RoboDK station: Doosan_M0609_SSM3_Experiment.rdk

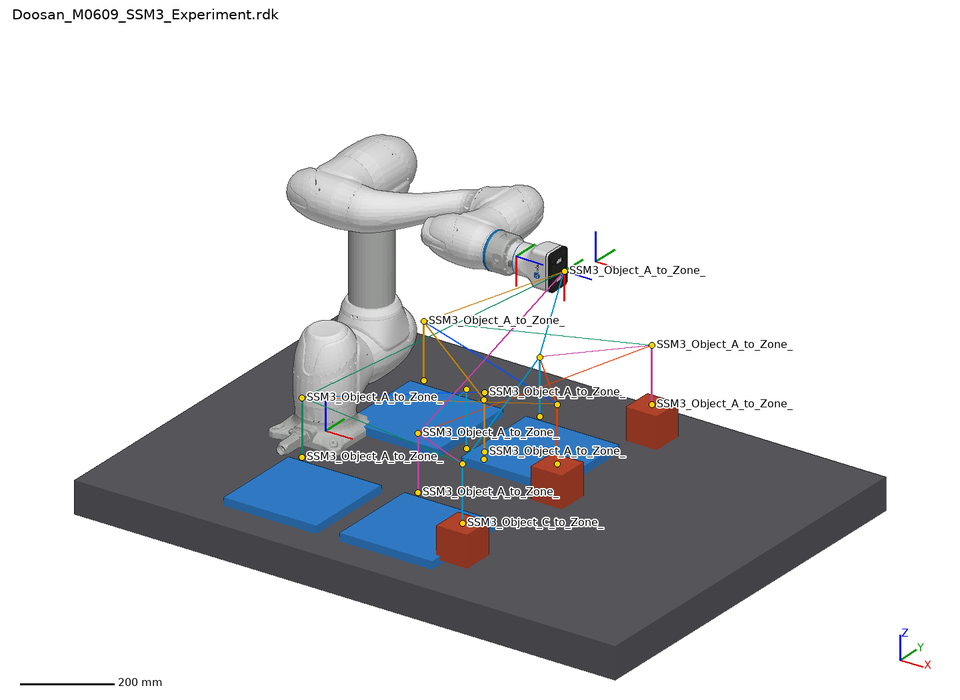
[picture v0: the station drawn from its stored meshes, robots at their saved joint values, targets as dots, program paths as lines]
Station Doosan_M0609_Pick_and_Place (saved by RoboDK 6.1.1). Poses are relative to the parent item; angles as X-Y-Z fixed-axis rotations.
  - frame Robot_Base at (0, 0, 0) mm
    - robot Doosan Robotics M0609 White: 6 axes, payload 6 kg, reach 900 mm, repeatability 0.03 mm, weight 27 kg
        modified DH rows (alpha deg, a mm, theta deg, d mm): 0, 0, 0, 135; -90, 0, -90, -6.207; 0, 411, -90, 0; -90, 0, 0, 368; 90, 0, 0, 0; -90, 0, 180, 121
        base shift (0, 0, 0) mm, rotated rx 0 ry 0 rz 180 deg
        joint limits [-360, -360, -150, -360, -360, -360] to [360, 360, 150, 360, 360, 360]; home [0, 0, 90, 0, 0, 0]; saved at [0, 0, 90, 0, 0, 0]
      - tool SSM3_Motion_TCP, TCP at (0, 0, 125) mm
      - frame OnRobot-2FG7-Gripper at (0, 0, 0) mm
        - robot OnRobot-2FG7-Gripper-Mechanism: 1 axes
            joint limits [0] to [55]; home [0]; saved at [49.5]
      - frame AUTO_Attach_TCP at (0, 0, 125) mm
  - frame TEST3 at (0, 1000, 0) mm
  - frame SSM3_Workcell at (0, 0, 0) mm
    - object SSM3_Table at (400, 0, -40) mm, size 1400 x 1000 x 80 mm, geometry from SSM3_Table.stl
    - object SSM3_Zone_A at (150, -300, 10) mm, size 240 x 240 x 20 mm, geometry from SSM3_Zone_A.stl
    - object SSM3_Zone_B at (450, -300, 10) mm, size 240 x 240 x 20 mm, geometry from SSM3_Zone_B.stl
    - object SSM3_Zone_C at (150, 150, 10) mm, size 240 x 240 x 20 mm, geometry from SSM3_Zone_C.stl
    - object SSM3_Zone_D at (450, 150, 10) mm, size 240 x 240 x 20 mm, geometry from SSM3_Zone_D.stl
    - target SSM3_Object_A_to_Zone_A_Home (Cartesian target) at (614, 6.21, 546) mm, rotated rx 0 ry 90 rz 0 deg; joints [0, 0, 90, 0, 0, 0] of Doosan Robotics M0609 White
    - target SSM3_Object_A_to_Zone_A_PickApproach (Cartesian target) at (440, -40, 230) mm, rotated rx 180 ry 0 rz 0 deg; joints [0, 0, 90, 0, 0, 0] of Doosan Robotics M0609 White
    - target SSM3_Object_A_to_Zone_A_Pick (Cartesian target) at (440, -40, 90) mm, rotated rx 180 ry 0 rz 0 deg; joints [0, 0, 90, 0, 0, 0] of Doosan Robotics M0609 White
    - target SSM3_Object_A_to_Zone_A_PlaceApproach (Cartesian target) at (150, -300, 240) mm, rotated rx 180 ry 0 rz 0 deg; joints [0, 0, 90, 0, 0, 0] of Doosan Robotics M0609 White
    - target SSM3_Object_A_to_Zone_A_Place (Cartesian target) at (150, -300, 100) mm, rotated rx 180 ry 0 rz 0 deg; joints [0, 0, 90, 0, 0, 0] of Doosan Robotics M0609 White
    - target SSM3_Object_A_to_Zone_B_Home (Cartesian target) at (614, 6.21, 546) mm, rotated rx 0 ry 90 rz 0 deg; joints [0, 0, 90, 0, 0, 0] of Doosan Robotics M0609 White
    - target SSM3_Object_A_to_Zone_B_PickApproach (Cartesian target) at (600, 350, 230) mm, rotated rx 180 ry 0 rz 0 deg; joints [0, 0, 90, 0, 0, 0] of Doosan Robotics M0609 White
    - target SSM3_Object_A_to_Zone_B_Pick (Cartesian target) at (600, 350, 90) mm, rotated rx 180 ry 0 rz 0 deg; joints [0, 0, 90, 0, 0, 0] of Doosan Robotics M0609 White
    - target SSM3_Object_A_to_Zone_B_PlaceApproach (Cartesian target) at (450, -300, 240) mm, rotated rx 180 ry 0 rz 0 deg; joints [0, 0, 90, 0, 0, 0] of Doosan Robotics M0609 White
    - target SSM3_Object_A_to_Zone_B_Place (Cartesian target) at (450, -300, 100) mm, rotated rx 180 ry 0 rz 0 deg; joints [0, 0, 90, 0, 0, 0] of Doosan Robotics M0609 White
    - target SSM3_Object_A_to_Zone_C_Home (Cartesian target) at (614, 6.21, 546) mm, rotated rx 0 ry 90 rz 0 deg; joints [0, 0, 90, 0, 0, 0] of Doosan Robotics M0609 White
    - target SSM3_Object_A_to_Zone_C_PickApproach (Cartesian target) at (600, 350, 230) mm, rotated rx 180 ry 0 rz 0 deg; joints [0, 0, 90, 0, 0, 0] of Doosan Robotics M0609 White
    - target SSM3_Object_A_to_Zone_C_Pick (Cartesian target) at (600, 350, 90) mm, rotated rx 180 ry 0 rz 0 deg; joints [0, 0, 90, 0, 0, 0] of Doosan Robotics M0609 White
    - target SSM3_Object_A_to_Zone_C_PlaceApproach (Cartesian target) at (150, 150, 240) mm, rotated rx 180 ry 0 rz 0 deg; joints [0, 0, 90, 0, 0, 0] of Doosan Robotics M0609 White
    - target SSM3_Object_A_to_Zone_C_Place (Cartesian target) at (150, 150, 100) mm, rotated rx 180 ry 0 rz 0 deg; joints [0, 0, 90, 0, 0, 0] of Doosan Robotics M0609 White
    - target SSM3_Object_A_to_Zone_D_Home (Cartesian target) at (614, 6.21, 546) mm, rotated rx 0 ry 90 rz 0 deg; joints [0, 0, 90, 0, 0, 0] of Doosan Robotics M0609 White
    - target SSM3_Object_A_to_Zone_D_PickApproach (Cartesian target) at (600, 350, 230) mm, rotated rx 180 ry 0 rz 0 deg; joints [0, 0, 90, 0, 0, 0] of Doosan Robotics M0609 White
    - target SSM3_Object_A_to_Zone_D_Pick (Cartesian target) at (600, 350, 90) mm, rotated rx 180 ry 0 rz 0 deg; joints [0, 0, 90, 0, 0, 0] of Doosan Robotics M0609 White
    - target SSM3_Object_A_to_Zone_D_PlaceApproach (Cartesian target) at (450, 150, 240) mm, rotated rx 180 ry 0 rz 0 deg; joints [0, 0, 90, 0, 0, 0] of Doosan Robotics M0609 White
    - target SSM3_Object_A_to_Zone_D_Place (Cartesian target) at (450, 150, 100) mm, rotated rx 180 ry 0 rz 0 deg; joints [0, 0, 90, 0, 0, 0] of Doosan Robotics M0609 White
    - target SSM3_Object_B_to_Zone_A_Home (Cartesian target) at (614, 6.21, 546) mm, rotated rx 0 ry 90 rz 0 deg; joints [0, 0, 90, 0, 0, 0] of Doosan Robotics M0609 White
    - target SSM3_Object_B_to_Zone_A_PickApproach (Cartesian target) at (600, 0, 230) mm, rotated rx 180 ry 0 rz 0 deg; joints [0, 0, 90, 0, 0, 0] of Doosan Robotics M0609 White
    - target SSM3_Object_B_to_Zone_A_Pick (Cartesian target) at (600, 0, 90) mm, rotated rx 180 ry 0 rz 0 deg; joints [0, 0, 90, 0, 0, 0] of Doosan Robotics M0609 White
    - target SSM3_Object_B_to_Zone_A_PlaceApproach (Cartesian target) at (150, -300, 240) mm, rotated rx 180 ry 0 rz 0 deg; joints [0, 0, 90, 0, 0, 0] of Doosan Robotics M0609 White
    - target SSM3_Object_B_to_Zone_A_Place (Cartesian target) at (150, -300, 100) mm, rotated rx 180 ry 0 rz 0 deg; joints [0, 0, 90, 0, 0, 0] of Doosan Robotics M0609 White
    - target SSM3_Object_B_to_Zone_B_Home (Cartesian target) at (614, 6.21, 546) mm, rotated rx 0 ry 90 rz 0 deg; joints [0, 0, 90, 0, 0, 0] of Doosan Robotics M0609 White
    - target SSM3_Object_B_to_Zone_B_PickApproach (Cartesian target) at (400, -50, 230) mm, rotated rx 180 ry 0 rz 0 deg; joints [0, 0, 90, 0, 0, 0] of Doosan Robotics M0609 White
    - target SSM3_Object_B_to_Zone_B_Pick (Cartesian target) at (400, -50, 90) mm, rotated rx 180 ry 0 rz 0 deg; joints [0, 0, 90, 0, 0, 0] of Doosan Robotics M0609 White
    - target SSM3_Object_B_to_Zone_B_PlaceApproach (Cartesian target) at (450, -300, 240) mm, rotated rx 180 ry 0 rz 0 deg; joints [0, 0, 90, 0, 0, 0] of Doosan Robotics M0609 White
    - target SSM3_Object_B_to_Zone_B_Place (Cartesian target) at (450, -300, 100) mm, rotated rx 180 ry 0 rz 0 deg; joints [0, 0, 90, 0, 0, 0] of Doosan Robotics M0609 White
    - target SSM3_Object_B_to_Zone_C_Home (Cartesian target) at (614, 6.21, 546) mm, rotated rx 0 ry 90 rz 0 deg; joints [0, 0, 90, 0, 0, 0] of Doosan Robotics M0609 White
    - target SSM3_Object_B_to_Zone_C_PickApproach (Cartesian target) at (600, 0, 230) mm, rotated rx 180 ry 0 rz 0 deg; joints [0, 0, 90, 0, 0, 0] of Doosan Robotics M0609 White
    - target SSM3_Object_B_to_Zone_C_Pick (Cartesian target) at (600, 0, 90) mm, rotated rx 180 ry 0 rz 0 deg; joints [0, 0, 90, 0, 0, 0] of Doosan Robotics M0609 White
    - target SSM3_Object_B_to_Zone_C_PlaceApproach (Cartesian target) at (150, 150, 240) mm, rotated rx 180 ry 0 rz 0 deg; joints [0, 0, 90, 0, 0, 0] of Doosan Robotics M0609 White
    - target SSM3_Object_B_to_Zone_C_Place (Cartesian target) at (150, 150, 100) mm, rotated rx 180 ry 0 rz 0 deg; joints [0, 0, 90, 0, 0, 0] of Doosan Robotics M0609 White
    - target SSM3_Object_B_to_Zone_D_Home (Cartesian target) at (614, 6.21, 546) mm, rotated rx 0 ry 90 rz 0 deg; joints [0, 0, 90, 0, 0, 0] of Doosan Robotics M0609 White
    - target SSM3_Object_B_to_Zone_D_PickApproach (Cartesian target) at (600, 0, 230) mm, rotated rx 180 ry 0 rz 0 deg; joints [0, 0, 90, 0, 0, 0] of Doosan Robotics M0609 White
    - target SSM3_Object_B_to_Zone_D_Pick (Cartesian target) at (600, 0, 90) mm, rotated rx 180 ry 0 rz 0 deg; joints [0, 0, 90, 0, 0, 0] of Doosan Robotics M0609 White
    - target SSM3_Object_B_to_Zone_D_PlaceApproach (Cartesian target) at (450, 150, 240) mm, rotated rx 180 ry 0 rz 0 deg; joints [0, 0, 90, 0, 0, 0] of Doosan Robotics M0609 White
    - target SSM3_Object_B_to_Zone_D_Place (Cartesian target) at (450, 150, 100) mm, rotated rx 180 ry 0 rz 0 deg; joints [0, 0, 90, 0, 0, 0] of Doosan Robotics M0609 White
    - target SSM3_Object_C_to_Zone_A_Home (Cartesian target) at (614, 6.21, 546) mm, rotated rx 0 ry 90 rz 0 deg; joints [0, 0, 90, 0, 0, 0] of Doosan Robotics M0609 White
    - target SSM3_Object_C_to_Zone_A_PickApproach (Cartesian target) at (600, -350, 230) mm, rotated rx 180 ry 0 rz 0 deg; joints [0, 0, 90, 0, 0, 0] of Doosan Robotics M0609 White
    - target SSM3_Object_C_to_Zone_A_Pick (Cartesian target) at (600, -350, 90) mm, rotated rx 180 ry 0 rz 0 deg; joints [0, 0, 90, 0, 0, 0] of Doosan Robotics M0609 White
    - target SSM3_Object_C_to_Zone_A_PlaceApproach (Cartesian target) at (150, -300, 240) mm, rotated rx 180 ry 0 rz 0 deg; joints [0, 0, 90, 0, 0, 0] of Doosan Robotics M0609 White
    - target SSM3_Object_C_to_Zone_A_Place (Cartesian target) at (150, -300, 100) mm, rotated rx 180 ry 0 rz 0 deg; joints [0, 0, 90, 0, 0, 0] of Doosan Robotics M0609 White
    - target SSM3_Object_C_to_Zone_B_Home (Cartesian target) at (614, 6.21, 546) mm, rotated rx 0 ry 90 rz 0 deg; joints [0, 0, 90, 0, 0, 0] of Doosan Robotics M0609 White
    - target SSM3_Object_C_to_Zone_B_PickApproach (Cartesian target) at (600, -350, 230) mm, rotated rx 180 ry 0 rz 0 deg; joints [0, 0, 90, 0, 0, 0] of Doosan Robotics M0609 White
    - target SSM3_Object_C_to_Zone_B_Pick (Cartesian target) at (600, -350, 90) mm, rotated rx 180 ry 0 rz 0 deg; joints [0, 0, 90, 0, 0, 0] of Doosan Robotics M0609 White
    - target SSM3_Object_C_to_Zone_B_PlaceApproach (Cartesian target) at (450, -300, 240) mm, rotated rx 180 ry 0 rz 0 deg; joints [0, 0, 90, 0, 0, 0] of Doosan Robotics M0609 White
    - target SSM3_Object_C_to_Zone_B_Place (Cartesian target) at (450, -300, 100) mm, rotated rx 180 ry 0 rz 0 deg; joints [0, 0, 90, 0, 0, 0] of Doosan Robotics M0609 White
    - target SSM3_Object_C_to_Zone_C_Home (Cartesian target) at (614, 6.21, 546) mm, rotated rx 0 ry 90 rz 0 deg; joints [0, 0, 90, 0, 0, 0] of Doosan Robotics M0609 White
    - target SSM3_Object_C_to_Zone_C_PickApproach (Cartesian target) at (460, -70, 230) mm, rotated rx 180 ry 0 rz 0 deg; joints [0, 0, 90, 0, 0, 0] of Doosan Robotics M0609 White
    - target SSM3_Object_C_to_Zone_C_Pick (Cartesian target) at (460, -70, 90) mm, rotated rx 180 ry 0 rz 0 deg; joints [0, 0, 90, 0, 0, 0] of Doosan Robotics M0609 White
    - target SSM3_Object_C_to_Zone_C_PlaceApproach (Cartesian target) at (150, 150, 240) mm, rotated rx 180 ry 0 rz 0 deg; joints [0, 0, 90, 0, 0, 0] of Doosan Robotics M0609 White
    - target SSM3_Object_C_to_Zone_C_Place (Cartesian target) at (150, 150, 100) mm, rotated rx 180 ry 0 rz 0 deg; joints [0, 0, 90, 0, 0, 0] of Doosan Robotics M0609 White
    - target SSM3_Object_C_to_Zone_D_Home (Cartesian target) at (614, 6.21, 546) mm, rotated rx 0 ry 90 rz 0 deg; joints [0, 0, 90, 0, 0, 0] of Doosan Robotics M0609 White
    - target SSM3_Object_C_to_Zone_D_PickApproach (Cartesian target) at (600, -350, 230) mm, rotated rx 180 ry 0 rz 0 deg; joints [0, 0, 90, 0, 0, 0] of Doosan Robotics M0609 White
    - target SSM3_Object_C_to_Zone_D_Pick (Cartesian target) at (600, -350, 90) mm, rotated rx 180 ry 0 rz 0 deg; joints [0, 0, 90, 0, 0, 0] of Doosan Robotics M0609 White
    - target SSM3_Object_C_to_Zone_D_PlaceApproach (Cartesian target) at (450, 150, 240) mm, rotated rx 180 ry 0 rz 0 deg; joints [0, 0, 90, 0, 0, 0] of Doosan Robotics M0609 White
    - target SSM3_Object_C_to_Zone_D_Place (Cartesian target) at (450, 150, 100) mm, rotated rx 180 ry 0 rz 0 deg; joints [0, 0, 90, 0, 0, 0] of Doosan Robotics M0609 White
    - object AUTO_Block at (600, 350, 50) mm, size 80 x 80 x 80 mm, geometry from AUTO_Block.stl
    - object SSM3_Object_B at (600, 0, 50) mm, size 80 x 80 x 80 mm, geometry from SSM3_Object_B.stl
    - object SSM3_Object_C at (600, -350, 50) mm, size 80 x 80 x 80 mm, geometry from SSM3_Object_C.stl
  - program PickPlace_Object_A_to_Zone_A (13 instructions, listed below)
  - program PickPlace_Object_A_to_Zone_B (13 instructions, listed below)
  - program PickPlace_Object_A_to_Zone_C (13 instructions, listed below)
  - program PickPlace_Object_A_to_Zone_D (13 instructions, listed below)
  - program PickPlace_Object_B_to_Zone_A (13 instructions, listed below)
  - program PickPlace_Object_B_to_Zone_B (13 instructions, listed below)
  - program PickPlace_Object_B_to_Zone_C (13 instructions, listed below)
  - program PickPlace_Object_B_to_Zone_D (13 instructions, listed below)
  - program PickPlace_Object_C_to_Zone_A (13 instructions, listed below)
  - program PickPlace_Object_C_to_Zone_B (13 instructions, listed below)
  - program PickPlace_Object_C_to_Zone_C (13 instructions, listed below)
  - program PickPlace_Object_C_to_Zone_D (13 instructions, listed below)
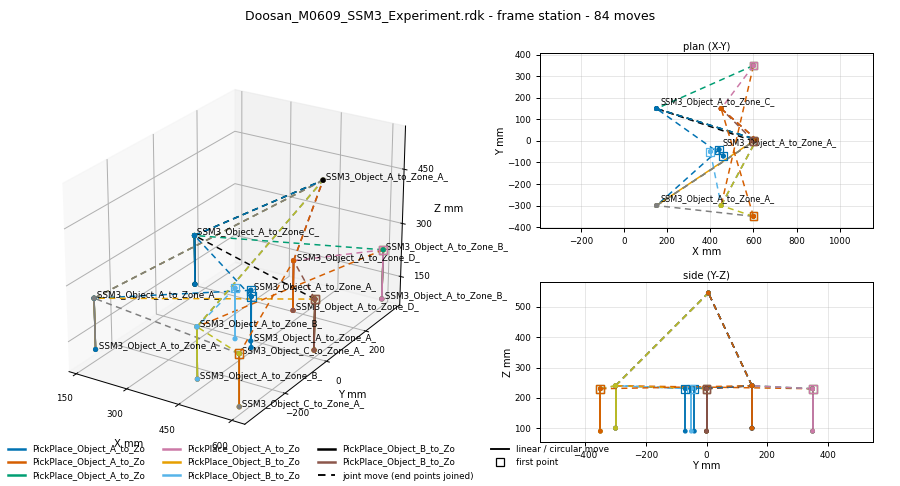
[picture p0: tool path of Doosan_M0609_SSM3_Experiment.rdk in frame station, 84 of 84 moves have a stored position in this frame; points joined in program order, loops and branches not executed]

--- program PickPlace_Object_A_to_Zone_A (robot Doosan Robotics M0609 White) ---
  Set Ref.: SSM3_Workcell
  Set Tool at (0, 0, 125) mm
  Set speed (60.0 mm/s)
  Set accel. (120.0 mm/s2)
  Set speed (10.0 deg/s)
  Set accel. (25.0 deg/s2)
  MoveJ (SSM3_Object_A_to_Zone_A_PickApproach)
  MoveL (SSM3_Object_A_to_Zone_A_Pick)
  MoveL (SSM3_Object_A_to_Zone_A_PickApproach)
  MoveJ (SSM3_Object_A_to_Zone_A_PlaceApproach)
  MoveL (SSM3_Object_A_to_Zone_A_Place)
  MoveL (SSM3_Object_A_to_Zone_A_PlaceApproach)
  MoveJ (SSM3_Object_A_to_Zone_A_Home)

--- program PickPlace_Object_A_to_Zone_B (robot Doosan Robotics M0609 White) ---
  Set Ref.: SSM3_Workcell
  Set Tool at (0, 0, 125) mm
  Set speed (60.0 mm/s)
  Set accel. (120.0 mm/s2)
  Set speed (10.0 deg/s)
  Set accel. (25.0 deg/s2)
  MoveJ (SSM3_Object_A_to_Zone_B_PickApproach)
  MoveL (SSM3_Object_A_to_Zone_B_Pick)
  MoveL (SSM3_Object_A_to_Zone_B_PickApproach)
  MoveJ (SSM3_Object_A_to_Zone_B_PlaceApproach)
  MoveL (SSM3_Object_A_to_Zone_B_Place)
  MoveL (SSM3_Object_A_to_Zone_B_PlaceApproach)
  MoveJ (SSM3_Object_A_to_Zone_B_Home)

--- program PickPlace_Object_A_to_Zone_C (robot Doosan Robotics M0609 White) ---
  Set Ref.: SSM3_Workcell
  Set Tool at (0, 0, 125) mm
  Set speed (60.0 mm/s)
  Set accel. (120.0 mm/s2)
  Set speed (10.0 deg/s)
  Set accel. (25.0 deg/s2)
  MoveJ (SSM3_Object_A_to_Zone_C_PickApproach)
  MoveL (SSM3_Object_A_to_Zone_C_Pick)
  MoveL (SSM3_Object_A_to_Zone_C_PickApproach)
  MoveJ (SSM3_Object_A_to_Zone_C_PlaceApproach)
  MoveL (SSM3_Object_A_to_Zone_C_Place)
  MoveL (SSM3_Object_A_to_Zone_C_PlaceApproach)
  MoveJ (SSM3_Object_A_to_Zone_C_Home)

--- program PickPlace_Object_A_to_Zone_D (robot Doosan Robotics M0609 White) ---
  Set Ref.: SSM3_Workcell
  Set Tool at (0, 0, 125) mm
  Set speed (60.0 mm/s)
  Set accel. (120.0 mm/s2)
  Set speed (10.0 deg/s)
  Set accel. (25.0 deg/s2)
  MoveJ (SSM3_Object_A_to_Zone_D_PickApproach)
  MoveL (SSM3_Object_A_to_Zone_D_Pick)
  MoveL (SSM3_Object_A_to_Zone_D_PickApproach)
  MoveJ (SSM3_Object_A_to_Zone_D_PlaceApproach)
  MoveL (SSM3_Object_A_to_Zone_D_Place)
  MoveL (SSM3_Object_A_to_Zone_D_PlaceApproach)
  MoveJ (SSM3_Object_A_to_Zone_D_Home)

--- program PickPlace_Object_B_to_Zone_A (robot Doosan Robotics M0609 White) ---
  Set Ref.: SSM3_Workcell
  Set Tool at (0, 0, 125) mm
  Set speed (60.0 mm/s)
  Set accel. (120.0 mm/s2)
  Set speed (10.0 deg/s)
  Set accel. (25.0 deg/s2)
  MoveJ (SSM3_Object_B_to_Zone_A_PickApproach)
  MoveL (SSM3_Object_B_to_Zone_A_Pick)
  MoveL (SSM3_Object_B_to_Zone_A_PickApproach)
  MoveJ (SSM3_Object_B_to_Zone_A_PlaceApproach)
  MoveL (SSM3_Object_B_to_Zone_A_Place)
  MoveL (SSM3_Object_B_to_Zone_A_PlaceApproach)
  MoveJ (SSM3_Object_B_to_Zone_A_Home)

--- program PickPlace_Object_B_to_Zone_B (robot Doosan Robotics M0609 White) ---
  Set Ref.: SSM3_Workcell
  Set Tool at (0, 0, 125) mm
  Set speed (60.0 mm/s)
  Set accel. (120.0 mm/s2)
  Set speed (10.0 deg/s)
  Set accel. (25.0 deg/s2)
  MoveJ (SSM3_Object_B_to_Zone_B_PickApproach)
  MoveL (SSM3_Object_B_to_Zone_B_Pick)
  MoveL (SSM3_Object_B_to_Zone_B_PickApproach)
  MoveJ (SSM3_Object_B_to_Zone_B_PlaceApproach)
  MoveL (SSM3_Object_B_to_Zone_B_Place)
  MoveL (SSM3_Object_B_to_Zone_B_PlaceApproach)
  MoveJ (SSM3_Object_B_to_Zone_B_Home)

--- program PickPlace_Object_B_to_Zone_C (robot Doosan Robotics M0609 White) ---
  Set Ref.: SSM3_Workcell
  Set Tool at (0, 0, 125) mm
  Set speed (60.0 mm/s)
  Set accel. (120.0 mm/s2)
  Set speed (10.0 deg/s)
  Set accel. (25.0 deg/s2)
  MoveJ (SSM3_Object_B_to_Zone_C_PickApproach)
  MoveL (SSM3_Object_B_to_Zone_C_Pick)
  MoveL (SSM3_Object_B_to_Zone_C_PickApproach)
  MoveJ (SSM3_Object_B_to_Zone_C_PlaceApproach)
  MoveL (SSM3_Object_B_to_Zone_C_Place)
  MoveL (SSM3_Object_B_to_Zone_C_PlaceApproach)
  MoveJ (SSM3_Object_B_to_Zone_C_Home)

--- program PickPlace_Object_B_to_Zone_D (robot Doosan Robotics M0609 White) ---
  Set Ref.: SSM3_Workcell
  Set Tool at (0, 0, 125) mm
  Set speed (60.0 mm/s)
  Set accel. (120.0 mm/s2)
  Set speed (10.0 deg/s)
  Set accel. (25.0 deg/s2)
  MoveJ (SSM3_Object_B_to_Zone_D_PickApproach)
  MoveL (SSM3_Object_B_to_Zone_D_Pick)
  MoveL (SSM3_Object_B_to_Zone_D_PickApproach)
  MoveJ (SSM3_Object_B_to_Zone_D_PlaceApproach)
  MoveL (SSM3_Object_B_to_Zone_D_Place)
  MoveL (SSM3_Object_B_to_Zone_D_PlaceApproach)
  MoveJ (SSM3_Object_B_to_Zone_D_Home)

--- program PickPlace_Object_C_to_Zone_A (robot Doosan Robotics M0609 White) ---
  Set Ref.: SSM3_Workcell
  Set Tool at (0, 0, 125) mm
  Set speed (60.0 mm/s)
  Set accel. (120.0 mm/s2)
  Set speed (10.0 deg/s)
  Set accel. (25.0 deg/s2)
  MoveJ (SSM3_Object_C_to_Zone_A_PickApproach)
  MoveL (SSM3_Object_C_to_Zone_A_Pick)
  MoveL (SSM3_Object_C_to_Zone_A_PickApproach)
  MoveJ (SSM3_Object_C_to_Zone_A_PlaceApproach)
  MoveL (SSM3_Object_C_to_Zone_A_Place)
  MoveL (SSM3_Object_C_to_Zone_A_PlaceApproach)
  MoveJ (SSM3_Object_C_to_Zone_A_Home)

--- program PickPlace_Object_C_to_Zone_B (robot Doosan Robotics M0609 White) ---
  Set Ref.: SSM3_Workcell
  Set Tool at (0, 0, 125) mm
  Set speed (60.0 mm/s)
  Set accel. (120.0 mm/s2)
  Set speed (10.0 deg/s)
  Set accel. (25.0 deg/s2)
  MoveJ (SSM3_Object_C_to_Zone_B_PickApproach)
  MoveL (SSM3_Object_C_to_Zone_B_Pick)
  MoveL (SSM3_Object_C_to_Zone_B_PickApproach)
  MoveJ (SSM3_Object_C_to_Zone_B_PlaceApproach)
  MoveL (SSM3_Object_C_to_Zone_B_Place)
  MoveL (SSM3_Object_C_to_Zone_B_PlaceApproach)
  MoveJ (SSM3_Object_C_to_Zone_B_Home)

--- program PickPlace_Object_C_to_Zone_C (robot Doosan Robotics M0609 White) ---
  Set Ref.: SSM3_Workcell
  Set Tool at (0, 0, 125) mm
  Set speed (60.0 mm/s)
  Set accel. (120.0 mm/s2)
  Set speed (10.0 deg/s)
  Set accel. (25.0 deg/s2)
  MoveJ (SSM3_Object_C_to_Zone_C_PickApproach)
  MoveL (SSM3_Object_C_to_Zone_C_Pick)
  MoveL (SSM3_Object_C_to_Zone_C_PickApproach)
  MoveJ (SSM3_Object_C_to_Zone_C_PlaceApproach)
  MoveL (SSM3_Object_C_to_Zone_C_Place)
  MoveL (SSM3_Object_C_to_Zone_C_PlaceApproach)
  MoveJ (SSM3_Object_C_to_Zone_C_Home)

--- program PickPlace_Object_C_to_Zone_D (robot Doosan Robotics M0609 White) ---
  Set Ref.: SSM3_Workcell
  Set Tool at (0, 0, 125) mm
  Set speed (60.0 mm/s)
  Set accel. (120.0 mm/s2)
  Set speed (10.0 deg/s)
  Set accel. (25.0 deg/s2)
  MoveJ (SSM3_Object_C_to_Zone_D_PickApproach)
  MoveL (SSM3_Object_C_to_Zone_D_Pick)
  MoveL (SSM3_Object_C_to_Zone_D_PickApproach)
  MoveJ (SSM3_Object_C_to_Zone_D_PlaceApproach)
  MoveL (SSM3_Object_C_to_Zone_D_Place)
  MoveL (SSM3_Object_C_to_Zone_D_PlaceApproach)
  MoveJ (SSM3_Object_C_to_Zone_D_Home)
